(* IEC 61131-3 sources: rules_plc/examples/simple, 1 file *)

(* ---- hello.st ---- *)
{external}
FUNCTION puts : DINT
    VAR_INPUT {ref}
        text : STRING;
    END_VAR
END_FUNCTION

PROGRAM hello
    VAR
        x: DINT;
    END_VAR
    puts('hello from rules_plc!$N');
END_PROGRAM
